Universal Robots URScript: T012_zai-org_GLM-4.7-FP8_edit_perf_rep1.urscript

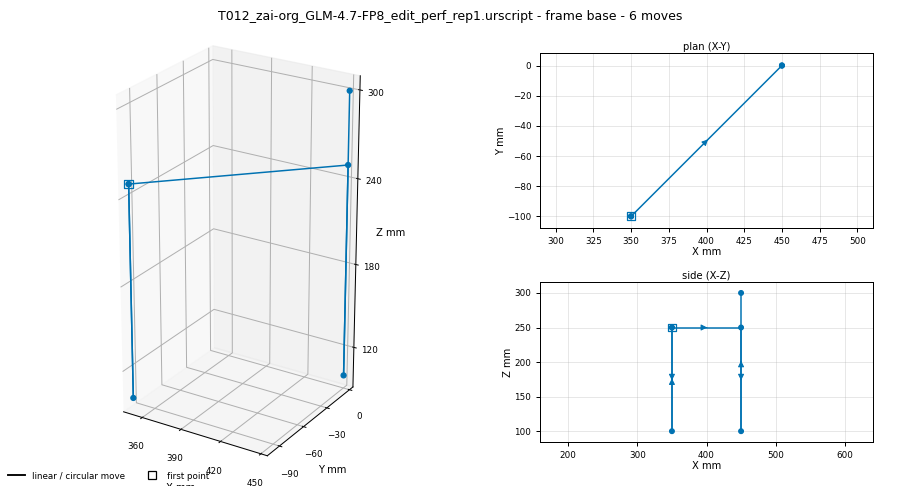
[picture p0: tool path of T012_zai-org_GLM-4.7-FP8_edit_perf_rep1.urscript in frame base, 6 of 8 moves have a stored position in this frame; points joined in program order, loops and branches not executed]
# Task: T012 — Collaborative spot welding — 3 points
# Optimized for faster cycle time
# Operating mode: collaborative | Max TCP speed: 0.250 m/s
# Robot: ur5e
#
# WARNING: This is auto-generated code for SIMULATION ONLY.
# Do NOT deploy to a physical robot without safety review.

def task_T012():
  # [0] E-Stop verify
  # E-Stop safety check (hardware-enforced on UR controller)
  if (get_digital_in(0) == True):
    popup("E-Stop active — aborting program.", error=True)
    halt
  end

  # [1] Home
  # Increased joint velocity and acceleration for faster repositioning
  movej([0.0000, -1.5708, 1.5708, -1.5708, -1.5708, 0.0000], a=2.0, v=2.0)

  # [2] Approach spot 1
  # Maximized TCP speed (0.25 m/s) and increased acceleration
  movel(p[0.350000, -0.100000, 0.250000, 0.0000, 3.1416, 0.0000], a=1.2, v=0.25, r=0.0)

  # [3] Descend to spot 1
  # Slightly increased descent speed for efficiency while maintaining precision
  movel(p[0.350000, -0.100000, 0.100000, 0.0000, 3.1416, 0.0000], a=0.5, v=0.10, r=0.0)

  # [4] Weld spot 1 ON
  # Welding arc ON (I=80A, wire=0.0m/min)
  set_digital_out(0, True)   # arc enable
  set_analog_out(0, 0.267)  # current (normalized)
  set_analog_out(1, 0.000)  # wire feed (normalized)

  # [5] Weld dwell
  sleep(0.5000)

  # [6] Weld spot 1 OFF
  # Welding arc OFF
  set_digital_out(0, False)
  set_analog_out(0, 0.0)
  set_analog_out(1, 0.0)

  # [7] Lift from spot 1
  # Increased speed and added blend radius (r=0.02) to smooth transition to next move
  movel(p[0.350000, -0.100000, 0.250000, 0.0000, 3.1416, 0.0000], a=1.2, v=0.25, r=0.02)

  # [8] Move to spot 2
  # Maximized TCP speed and acceleration
  movel(p[0.450000, 0.000000, 0.250000, 0.0000, 3.1416, 0.0000], a=1.2, v=0.25, r=0.0)

  # [9] Descend to spot 2
  # Slightly increased descent speed
  movel(p[0.450000, 0.000000, 0.100000, 0.0000, 3.1416, 0.0000], a=0.5, v=0.10, r=0.0)

  # [10] Weld spot 2 ON
  # Welding arc ON (I=80A, wire=0.0m/min)
  set_digital_out(0, True)   # arc enable
  set_analog_out(0, 0.267)  # current (normalized)
  set_analog_out(1, 0.000)  # wire feed (normalized)

  # [11] Weld dwell
  sleep(0.5000)

  # [12] Weld spot 2 OFF
  # Welding arc OFF
  set_digital_out(0, False)
  set_analog_out(0, 0.0)
  set_analog_out(1, 0.0)

  # [13] Retract
  # Increased speed and added blend radius (r=0.02) to smooth transition to Home
  movel(p[0.450000, 0.000000, 0.300000, 0.0000, 3.1416, 0.0000], a=1.2, v=0.25, r=0.02)

  # [14] Return home
  # Increased joint velocity and acceleration
  movej([0.0000, -1.5708, 1.5708, -1.5708, -1.5708, 0.0000], a=2.0, v=2.0)

end

# Entry point
task_T012()
